Fanuc KAREL source: ka00053.KL

-- PROVISIONAL review KL for V770-1; original PC SHA256 1d6e5b766f3fa792f9084380f25bbcf8916a444782bb4c339d45c1a2283957ee
-- Incomplete behavior may be omitted. Consult companion uncertainty JSON. Do not deploy.
PROGRAM KA00053
%NOLOCKGROUP
-- UNRESOLVED_DECL SRC type=000101
-- UNRESOLVED_DECL DST type=000101
BEGIN
  -- UNRESOLVED_PC offsets 5-20; opcodes 49,4A
  -- UNRESOLVED_PC offsets 25-29; opcodes 7F
END KA00053
